// TIA Portal V21 export
// export: Created 2026-08-21T20:18:50.9416653Z, ExportSetting None, DisplayName Totally Integrated Automation Portal, DisplayVersion V21, DisplayName STEP 7 Professional, DisplayVersion V21, DisplayName STEP 7 Safety, DisplayVersion V21, DisplayName Tech WebApplication, DisplayVersion V21, DisplayName WinCC Basic/Comfort/Advanced, DisplayVersion V21, DisplayName WinCC Professional, DisplayVersion V21, DisplayName WinCC Unified, DisplayVersion V21
FUNCTION "LIT100" : Void   // FC6, FBD
{ S7_Optimized_Access := 'TRUE' }
// stored: SetENOAutomatically false
BEGIN

REGION Network 1: Tank level
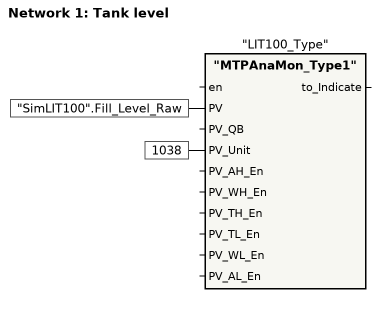
   "LIT100_Type"(PV := "SimLIT100".Fill_Level_Raw, PV_Unit := 1038);   // "MTPAnaMon_Type1"
END_REGION
END_FUNCTION
